// TIA Portal V19 export
TYPE "EM_Output"
   STRUCT
      ModeMan : Bool;
      ModeAuto : Bool;
      ModeMaint : Bool;
      ModeConflict : Bool;   // MÃ¡s de un modo solicitado a la vez
      Idle : Bool;
      Running : Bool;
      Completed : Bool;
      Holding : Bool;
      Held : Bool;
      Stopping : Bool;
      Stopped : Bool;
      Aborting : Bool;
      Aborted : Bool;
      Fault : Bool;
      State : Int;   // 0=Idle 1=Running 2=Completed 3=Holding 4=Held 5=Stopping 6=Stopped 7=Aborting 8=Aborted
      FaultCode : Int;   // 0=Sin fallo 1=ParÃ¡metros invÃ¡lidos 2=Sensor de temperatura invÃ¡lido 3=Timeout de temperatura 4=VÃ¡lvula no abre 5=Alarma del CM 6=VÃ¡lvula no cierra 7=ConcSMMV fuera de rango (0..100)
   END_STRUCT;
END_TYPE
